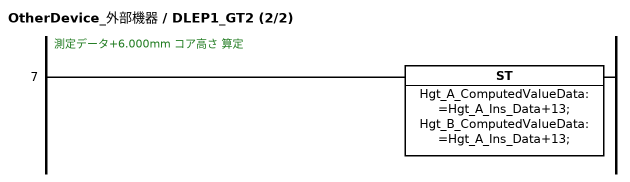
(* [picture p96: OtherDevice_外部機器 / DLEP1_GT2, rungs 7-7] *)
(* Rung 7: 測定データ+6.000mm コア高さ 算定 *)
Hgt_A_ComputedValueData:=Hgt_A_Ins_Data+13;
Hgt_B_ComputedValueData:=Hgt_A_Ins_Data+13;

(* Section FH_5552_10: ladder, written here as Structured Text *)

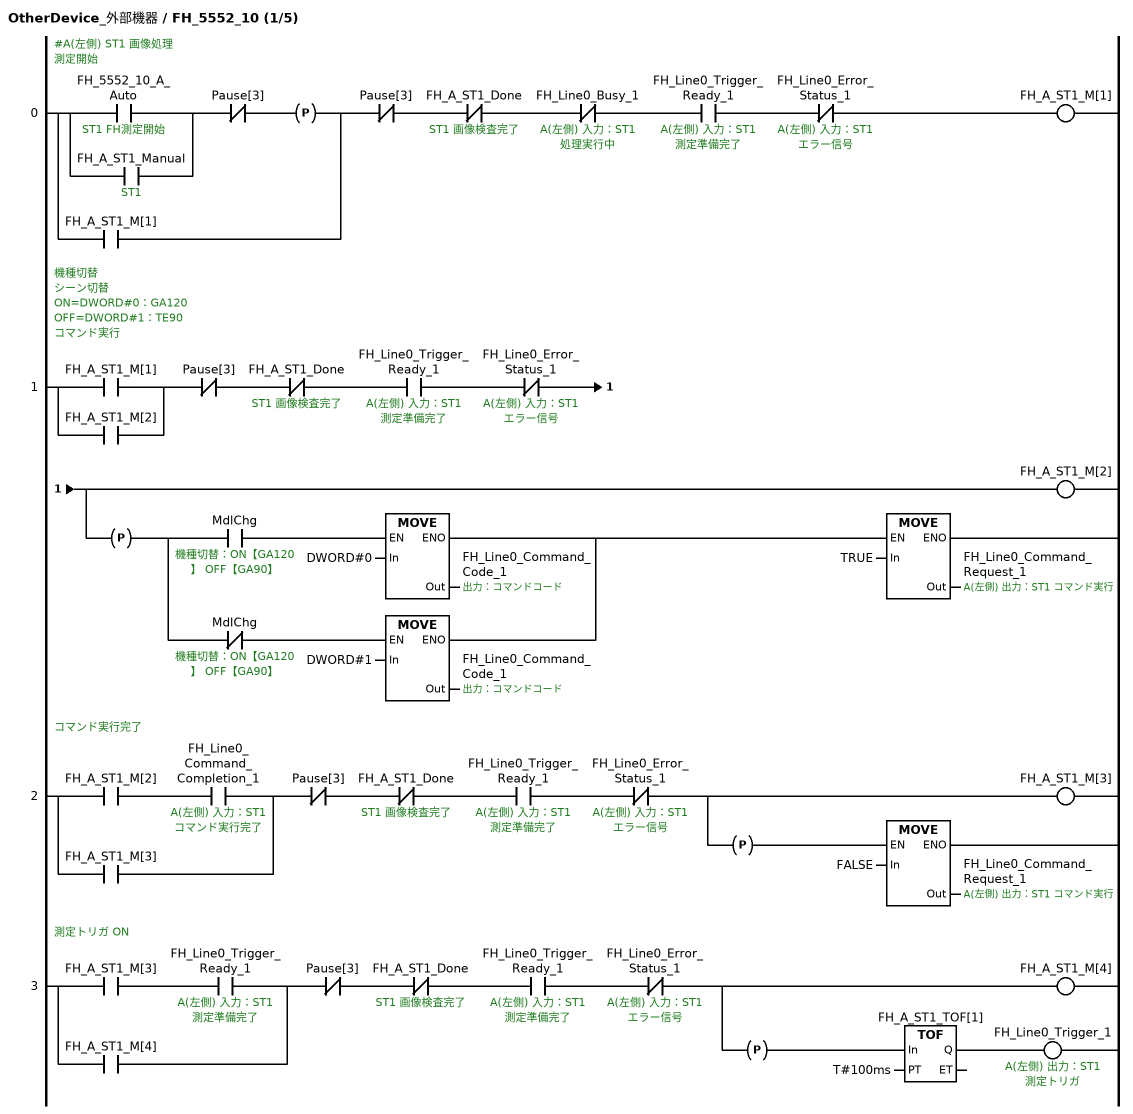
(* Rung 0: #A(左側) ST1 画像処理 / 測定開始 *)
_e25(CLK := (FH_5552_10_A_Auto OR FH_A_ST1_Manual) AND NOT Pause[3]);
FH_A_ST1_M[1] := (_e25.Q OR FH_A_ST1_M[1]) AND NOT Pause[3] AND NOT FH_A_ST1_Done AND NOT FH_Line0_Busy_1 AND FH_Line0_Trigger_Ready_1 AND NOT FH_Line0_Error_Status_1;
(* Rung 1: 機種切替 / シーン切替 / ON=DWORD#0：GA120 / OFF=DWORD#1：TE90 / コマンド実行 *)
_p26 := (FH_A_ST1_M[1] OR FH_A_ST1_M[2]) AND NOT Pause[3] AND NOT FH_A_ST1_Done AND FH_Line0_Trigger_Ready_1 AND NOT FH_Line0_Error_Status_1;
FH_A_ST1_M[2] := _p26;
_e27(CLK := _p26);
IF _e27.Q AND MdlChg THEN FH_Line0_Command_Code_1 := DWORD#0; END_IF;
IF _e27.Q AND NOT MdlChg THEN FH_Line0_Command_Code_1 := DWORD#1; END_IF;
IF _e27.Q AND (MdlChg OR NOT MdlChg) THEN FH_Line0_Command_Request_1 := TRUE; END_IF;
(* Rung 2: コマンド実行完了 *)
_p28 := ((FH_A_ST1_M[2] AND FH_Line0_Command_Completion_1) OR FH_A_ST1_M[3]) AND NOT Pause[3] AND NOT FH_A_ST1_Done AND FH_Line0_Trigger_Ready_1 AND NOT FH_Line0_Error_Status_1;
FH_A_ST1_M[3] := _p28;
_e29(CLK := _p28);
IF _e29.Q THEN FH_Line0_Command_Request_1 := FALSE; END_IF;
(* Rung 3: 測定トリガ ON *)
_p30 := ((FH_A_ST1_M[3] AND FH_Line0_Trigger_Ready_1) OR FH_A_ST1_M[4]) AND NOT Pause[3] AND NOT FH_A_ST1_Done AND FH_Line0_Trigger_Ready_1 AND NOT FH_Line0_Error_Status_1;
FH_A_ST1_M[4] := _p30;
_e31(CLK := _p30);
FH_A_ST1_TOF[1](In := _e31.Q, PT := T#100ms);
FH_Line0_Trigger_1 := FH_A_ST1_TOF[1].Q;

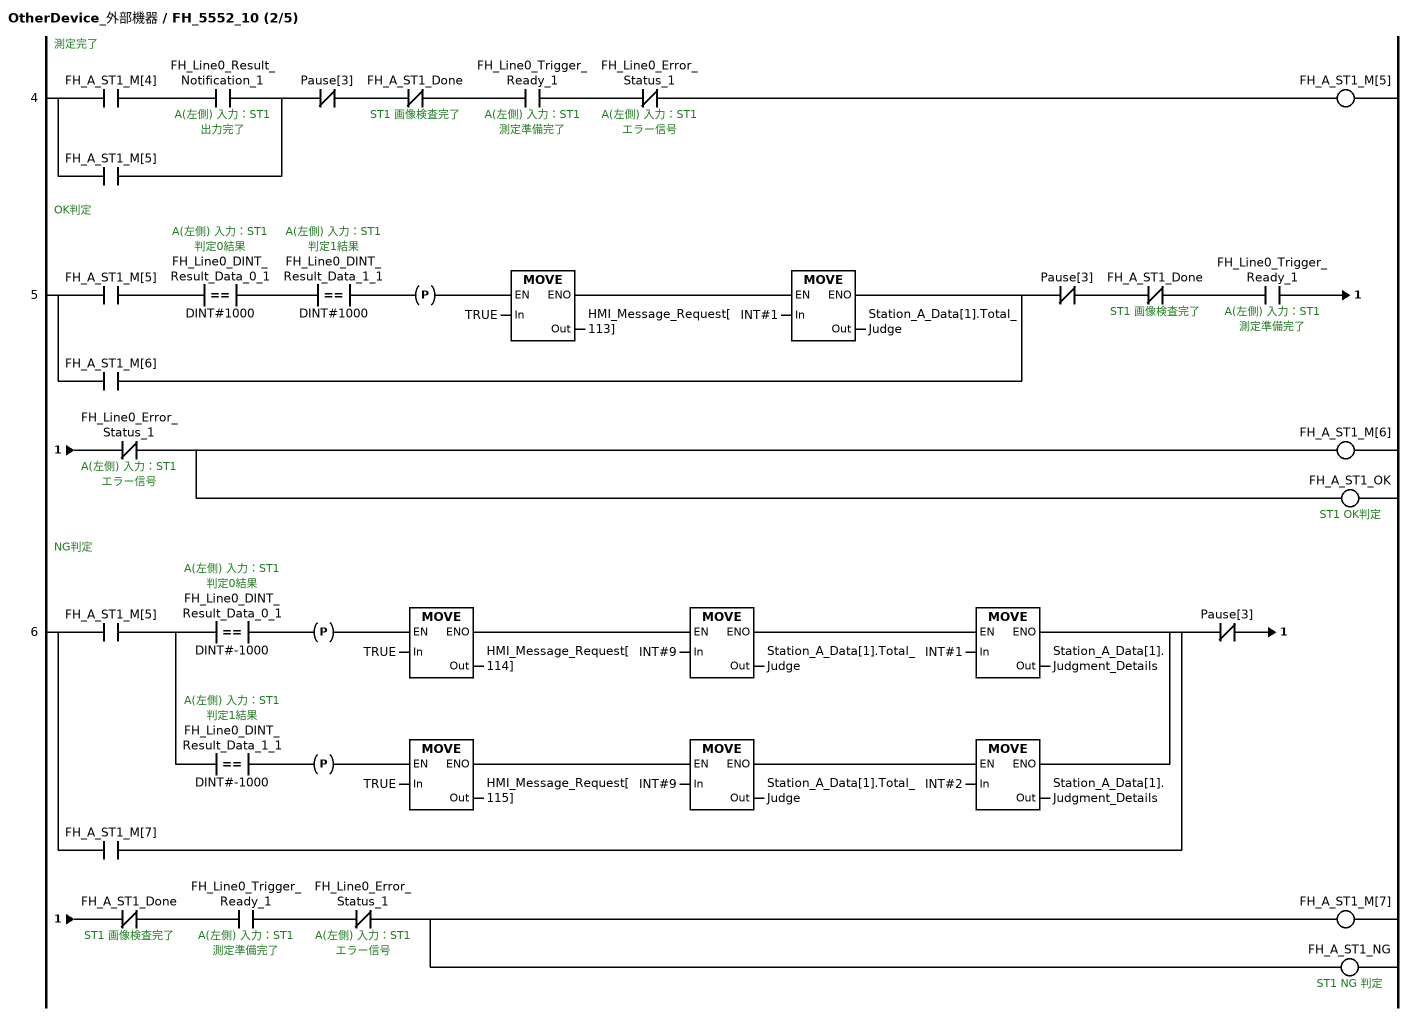
(* Rung 4: 測定完了 *)
FH_A_ST1_M[5] := ((FH_A_ST1_M[4] AND FH_Line0_Result_Notification_1) OR FH_A_ST1_M[5]) AND NOT Pause[3] AND NOT FH_A_ST1_Done AND FH_Line0_Trigger_Ready_1 AND NOT FH_Line0_Error_Status_1;
(* Rung 5: OK判定 *)
_e32(CLK := FH_A_ST1_M[5] AND (FH_Line0_DINT_Result_Data_0_1 = DINT#1000) AND (FH_Line0_DINT_Result_Data_1_1 = DINT#1000));
IF _e32.Q THEN
    HMI_Message_Request[113] := TRUE;
    Station_A_Data[1].Total_Judge := INT#1;
END_IF;
_p33 := (_e32.Q OR FH_A_ST1_M[6]) AND NOT Pause[3] AND NOT FH_A_ST1_Done AND FH_Line0_Trigger_Ready_1 AND NOT FH_Line0_Error_Status_1;
FH_A_ST1_M[6] := _p33;
FH_A_ST1_OK := _p33;
(* Rung 6: NG判定 *)
_e34(CLK := FH_A_ST1_M[5] AND (FH_Line0_DINT_Result_Data_0_1 = (DINT#-1000)));
IF _e34.Q THEN
    HMI_Message_Request[114] := TRUE;
    Station_A_Data[1].Total_Judge := INT#9;
    Station_A_Data[1].Judgment_Details := INT#1;
END_IF;
_e35(CLK := FH_A_ST1_M[5] AND (FH_Line0_DINT_Result_Data_1_1 = (DINT#-1000)));
IF _e35.Q THEN
    HMI_Message_Request[115] := TRUE;
    Station_A_Data[1].Total_Judge := INT#9;
    Station_A_Data[1].Judgment_Details := INT#2;
END_IF;
_p36 := (_e34.Q OR _e35.Q OR FH_A_ST1_M[7]) AND NOT Pause[3] AND NOT FH_A_ST1_Done AND FH_Line0_Trigger_Ready_1 AND NOT FH_Line0_Error_Status_1;
FH_A_ST1_M[7] := _p36;
FH_A_ST1_NG := _p36;

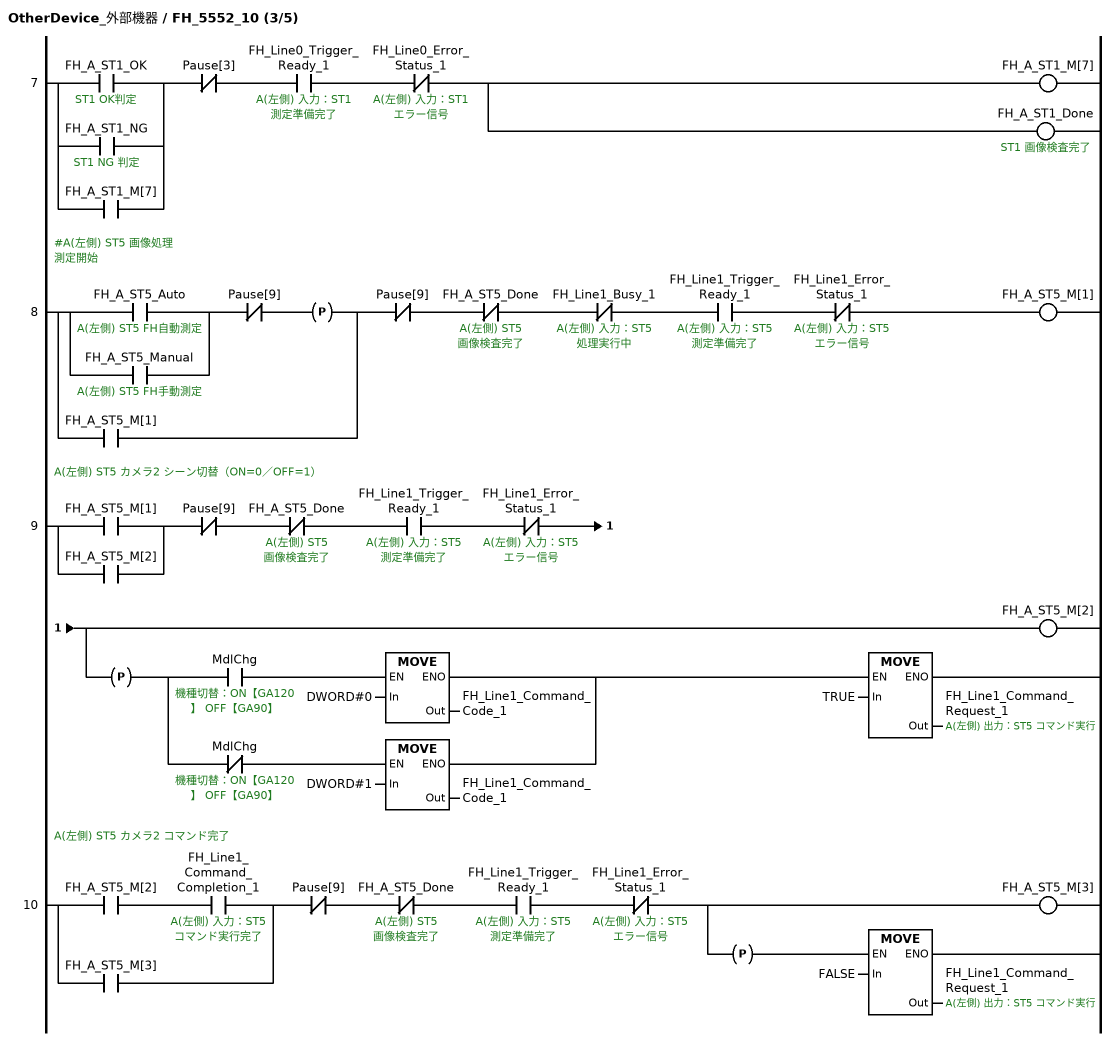
(* Rung 7 *)
_p37 := (FH_A_ST1_OK OR FH_A_ST1_NG OR FH_A_ST1_M[7]) AND NOT Pause[3] AND FH_Line0_Trigger_Ready_1 AND NOT FH_Line0_Error_Status_1;
FH_A_ST1_M[7] := _p37;
FH_A_ST1_Done := _p37;
(* Rung 8: #A(左側) ST5 画像処理 / 測定開始 *)
_e38(CLK := (FH_A_ST5_Auto OR FH_A_ST5_Manual) AND NOT Pause[9]);
FH_A_ST5_M[1] := (_e38.Q OR FH_A_ST5_M[1]) AND NOT Pause[9] AND NOT FH_A_ST5_Done AND NOT FH_Line1_Busy_1 AND FH_Line1_Trigger_Ready_1 AND NOT FH_Line1_Error_Status_1;
(* Rung 9: A(左側) ST5 カメラ2 シーン切替（ON=0／OFF=1） *)
_p39 := (FH_A_ST5_M[1] OR FH_A_ST5_M[2]) AND NOT Pause[9] AND NOT FH_A_ST5_Done AND FH_Line1_Trigger_Ready_1 AND NOT FH_Line1_Error_Status_1;
FH_A_ST5_M[2] := _p39;
_e40(CLK := _p39);
IF _e40.Q AND MdlChg THEN FH_Line1_Command_Code_1 := DWORD#0; END_IF;
IF _e40.Q AND NOT MdlChg THEN FH_Line1_Command_Code_1 := DWORD#1; END_IF;
IF _e40.Q AND (MdlChg OR NOT MdlChg) THEN FH_Line1_Command_Request_1 := TRUE; END_IF;
(* Rung 10: A(左側) ST5 カメラ2 コマンド完了 *)
_p41 := ((FH_A_ST5_M[2] AND FH_Line1_Command_Completion_1) OR FH_A_ST5_M[3]) AND NOT Pause[9] AND NOT FH_A_ST5_Done AND FH_Line1_Trigger_Ready_1 AND NOT FH_Line1_Error_Status_1;
FH_A_ST5_M[3] := _p41;
_e42(CLK := _p41);
IF _e42.Q THEN FH_Line1_Command_Request_1 := FALSE; END_IF;

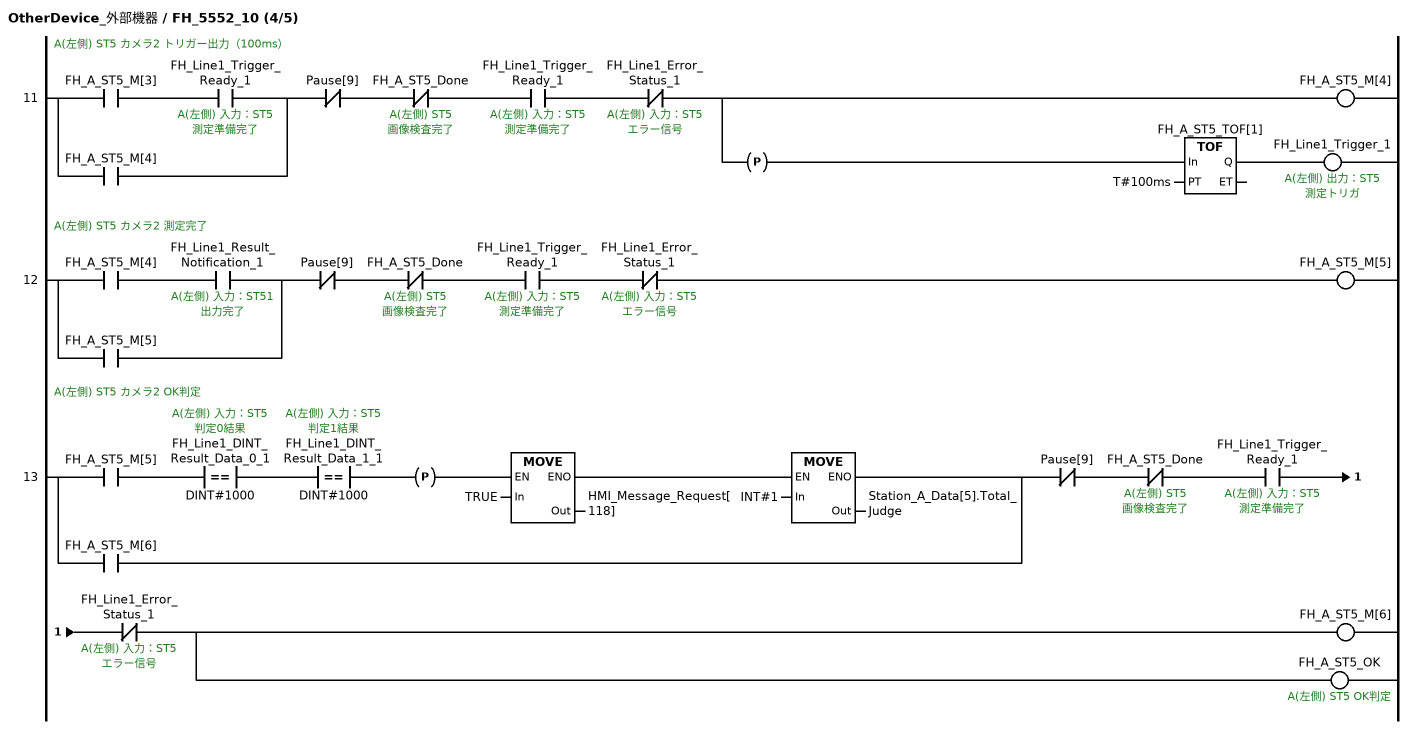
(* Rung 11: A(左側) ST5 カメラ2 トリガー出力（100ms） *)
_p43 := ((FH_A_ST5_M[3] AND FH_Line1_Trigger_Ready_1) OR FH_A_ST5_M[4]) AND NOT Pause[9] AND NOT FH_A_ST5_Done AND FH_Line1_Trigger_Ready_1 AND NOT FH_Line1_Error_Status_1;
FH_A_ST5_M[4] := _p43;
_e44(CLK := _p43);
FH_A_ST5_TOF[1](In := _e44.Q, PT := T#100ms);
FH_Line1_Trigger_1 := FH_A_ST5_TOF[1].Q;
(* Rung 12: A(左側) ST5 カメラ2 測定完了 *)
FH_A_ST5_M[5] := ((FH_A_ST5_M[4] AND FH_Line1_Result_Notification_1) OR FH_A_ST5_M[5]) AND NOT Pause[9] AND NOT FH_A_ST5_Done AND FH_Line1_Trigger_Ready_1 AND NOT FH_Line1_Error_Status_1;
(* Rung 13: A(左側) ST5 カメラ2 OK判定 *)
_e45(CLK := FH_A_ST5_M[5] AND (FH_Line1_DINT_Result_Data_0_1 = DINT#1000) AND (FH_Line1_DINT_Result_Data_1_1 = DINT#1000));
IF _e45.Q THEN
    HMI_Message_Request[118] := TRUE;
    Station_A_Data[5].Total_Judge := INT#1;
END_IF;
_p46 := (_e45.Q OR FH_A_ST5_M[6]) AND NOT Pause[9] AND NOT FH_A_ST5_Done AND FH_Line1_Trigger_Ready_1 AND NOT FH_Line1_Error_Status_1;
FH_A_ST5_M[6] := _p46;
FH_A_ST5_OK := _p46;

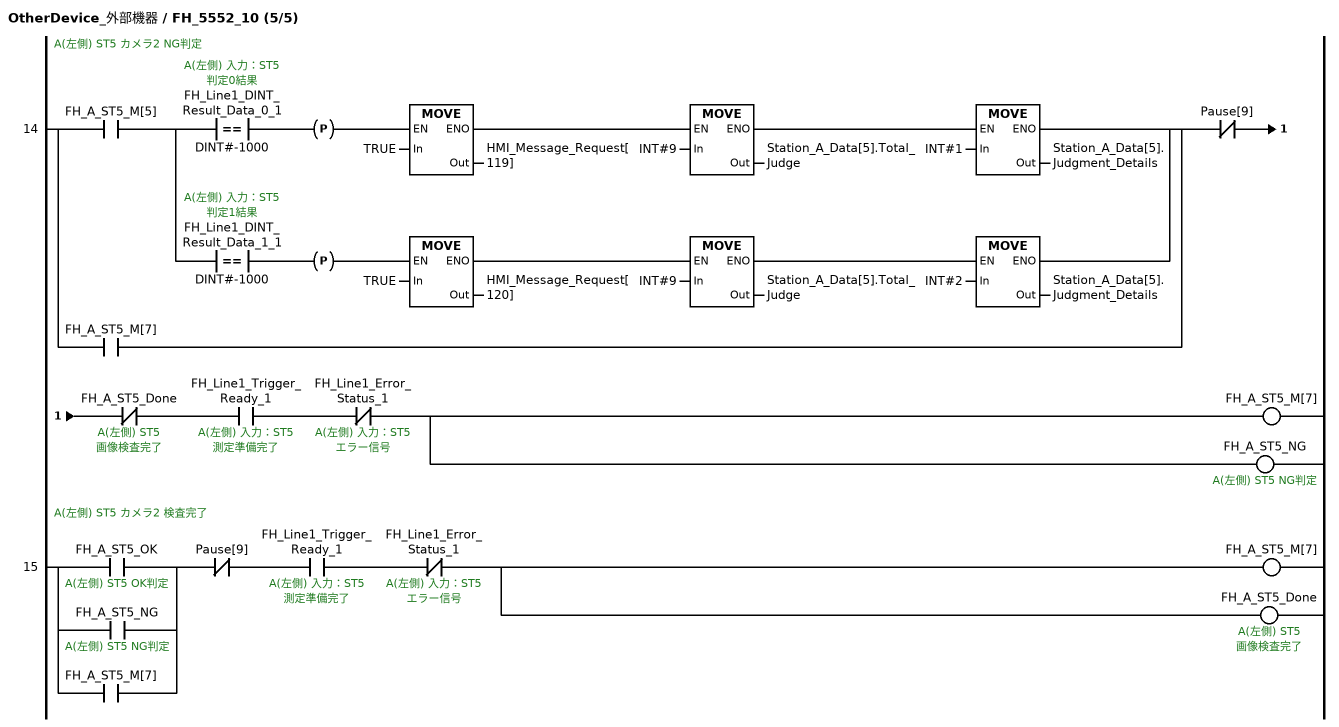
(* Rung 14: A(左側) ST5 カメラ2 NG判定 *)
_e47(CLK := FH_A_ST5_M[5] AND (FH_Line1_DINT_Result_Data_0_1 = (DINT#-1000)));
IF _e47.Q THEN
    HMI_Message_Request[119] := TRUE;
    Station_A_Data[5].Total_Judge := INT#9;
    Station_A_Data[5].Judgment_Details := INT#1;
END_IF;
_e48(CLK := FH_A_ST5_M[5] AND (FH_Line1_DINT_Result_Data_1_1 = (DINT#-1000)));
IF _e48.Q THEN
    HMI_Message_Request[120] := TRUE;
    Station_A_Data[5].Total_Judge := INT#9;
    Station_A_Data[5].Judgment_Details := INT#2;
END_IF;
_p49 := (_e47.Q OR _e48.Q OR FH_A_ST5_M[7]) AND NOT Pause[9] AND NOT FH_A_ST5_Done AND FH_Line1_Trigger_Ready_1 AND NOT FH_Line1_Error_Status_1;
FH_A_ST5_M[7] := _p49;
FH_A_ST5_NG := _p49;
(* Rung 15: A(左側) ST5 カメラ2 検査完了 *)
_p50 := (FH_A_ST5_OK OR FH_A_ST5_NG OR FH_A_ST5_M[7]) AND NOT Pause[9] AND FH_Line1_Trigger_Ready_1 AND NOT FH_Line1_Error_Status_1;
FH_A_ST5_M[7] := _p50;
FH_A_ST5_Done := _p50;

(* Section CV2A_KED: ladder, written here as Structured Text *)

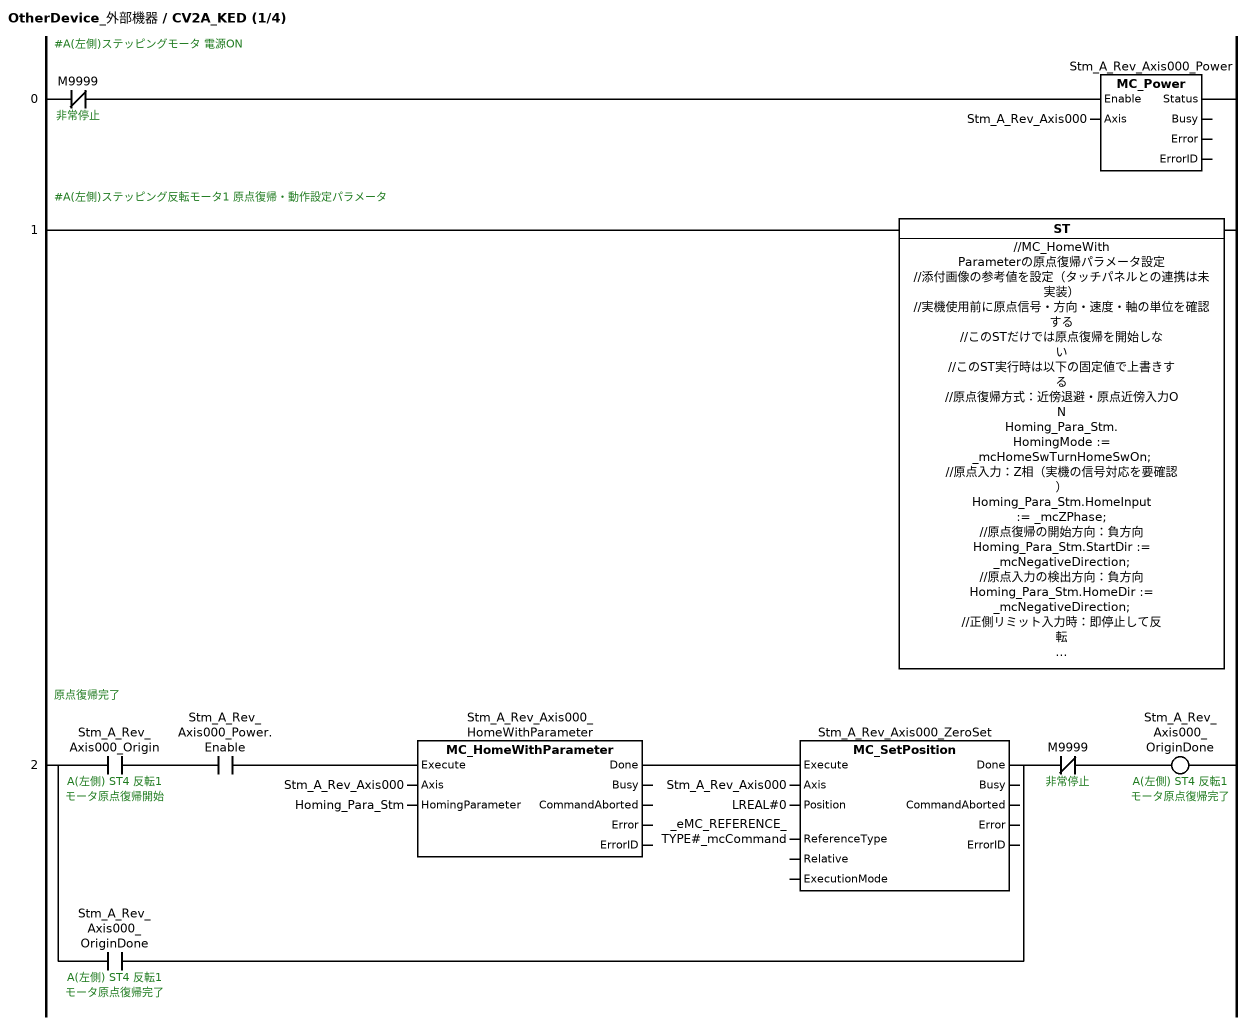
(* Rung 0: #A(左側)ステッピングモータ 電源ON *)
Stm_A_Rev_Axis000_Power(Enable := NOT M9999, Axis := Stm_A_Rev_Axis000);
(* Rung 1: #A(左側)ステッピング反転モータ1 原点復帰・動作設定パラメータ *)
//MC_HomeWithParameterの原点復帰パラメータ設定
//添付画像の参考値を設定（タッチパネルとの連携は未実装）
//実機使用前に原点信号・方向・速度・軸の単位を確認する
//このSTだけでは原点復帰を開始しない
//このST実行時は以下の固定値で上書きする

//原点復帰方式：近傍退避・原点近傍入力ON
Homing_Para_Stm.HomingMode := _mcHomeSwTurnHomeSwOn;
//原点入力：Z相（実機の信号対応を要確認）
Homing_Para_Stm.HomeInput := _mcZPhase;
//原点復帰の開始方向：負方向
Homing_Para_Stm.StartDir := _mcNegativeDirection;
//原点入力の検出方向：負方向
Homing_Para_Stm.HomeDir := _mcNegativeDirection;
//正側リミット入力時：即停止して反転
Homing_Para_Stm.PosiLmtMode := _mcRevImmediateStop;
//負側リミット入力時：即停止して反転
Homing_Para_Stm.NegaLmtMode := _mcRevImmediateStop;

//原点復帰速度 [指令単位/s]
Homing_Para_Stm.Vel := LREAL#40;
//原点近傍での接近速度 [指令単位/s]
Homing_Para_Stm.ApproachVel := LREAL#1;
//原点復帰の加速度 [指令単位/s^2]
Homing_Para_Stm.Acc := LREAL#100;
//原点復帰の減速度 [指令単位/s^2]
Homing_Para_Stm.Dec := LREAL#200;
//ジャーク [指令単位/s^3]：0はジャーク制御なし
Homing_Para_Stm.Jerk := LREAL#0;

//原点入力マスク距離 [指令単位]：今回の方式では未使用
Homing_Para_Stm.Mask := LREAL#0;
//原点確定後の現在位置 [指令単位]
Homing_Para_Stm.Offset := LREAL#0;
//押当て時間 [ms]：今回の方式では未使用
Homing_Para_Stm.PushTime := UINT#0;
//原点検出後の補正移動量 [指令単位]：0は補正移動なし
Homing_Para_Stm.Compensation := LREAL#0;
//原点補正移動時の速度 [指令単位/s]
Homing_Para_Stm.CompensationVel := LREAL#10;
(* Rung 2: 原点復帰完了 *)
Stm_A_Rev_Axis000_HomeWithParameter(Execute := Stm_A_Rev_Axis000_Origin AND Stm_A_Rev_Axis000_Power.Enable, Axis := Stm_A_Rev_Axis000, HomingParameter := Homing_Para_Stm);
Stm_A_Rev_Axis000_ZeroSet(Execute := Stm_A_Rev_Axis000_HomeWithParameter.Done, Axis := Stm_A_Rev_Axis000, Position := LREAL#0, ReferenceType := _eMC_REFERENCE_TYPE#_mcCommand);
Stm_A_Rev_Axis000_OriginDone := (Stm_A_Rev_Axis000_ZeroSet.Done OR Stm_A_Rev_Axis000_OriginDone) AND NOT M9999;

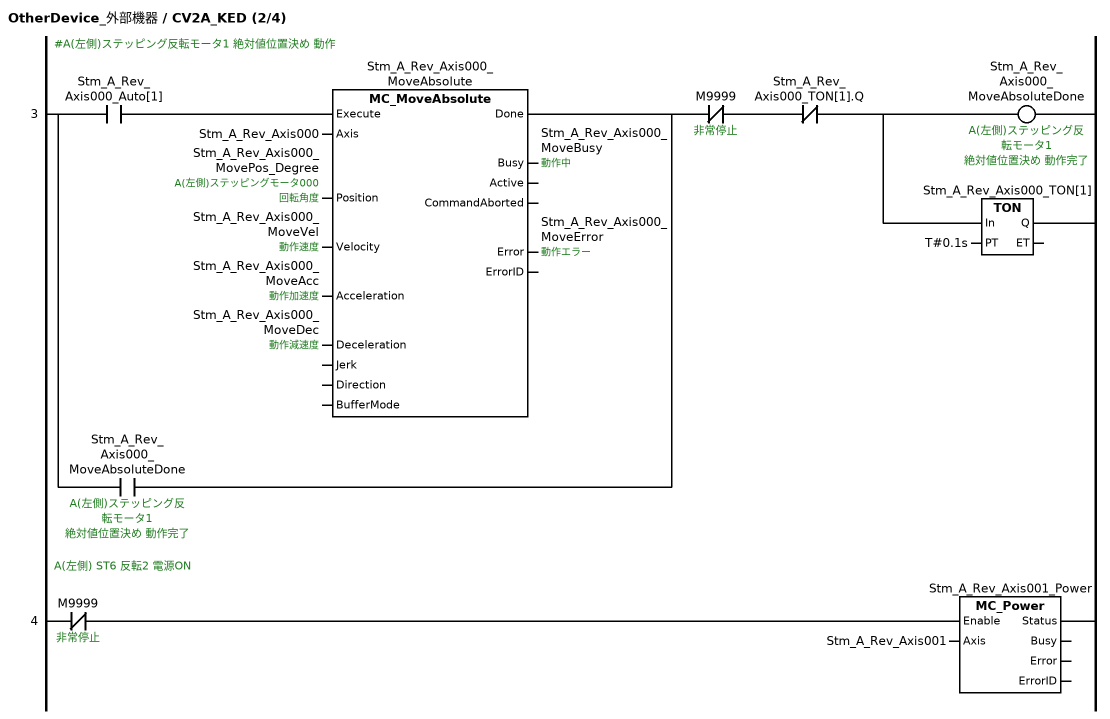
(* Rung 3: #A(左側)ステッピング反転モータ1 絶対値位置決め 動作 *)
Stm_A_Rev_Axis000_MoveAbsolute(Execute := Stm_A_Rev_Axis000_Auto[1], Axis := Stm_A_Rev_Axis000, Position := Stm_A_Rev_Axis000_MovePos_Degree, Velocity := Stm_A_Rev_Axis000_MoveVel, Acceleration := Stm_A_Rev_Axis000_MoveAcc, Deceleration := Stm_A_Rev_Axis000_MoveDec, Busy => Stm_A_Rev_Axis000_MoveBusy, Error => Stm_A_Rev_Axis000_MoveError);
_p51 := (Stm_A_Rev_Axis000_MoveAbsolute.Done OR Stm_A_Rev_Axis000_MoveAbsoluteDone) AND NOT M9999 AND NOT Stm_A_Rev_Axis000_TON[1].Q;
Stm_A_Rev_Axis000_MoveAbsoluteDone := _p51;
Stm_A_Rev_Axis000_TON[1](In := _p51, PT := T#0.1s);
(* Rung 4: A(左側) ST6 反転2 電源ON *)
Stm_A_Rev_Axis001_Power(Enable := NOT M9999, Axis := Stm_A_Rev_Axis001);

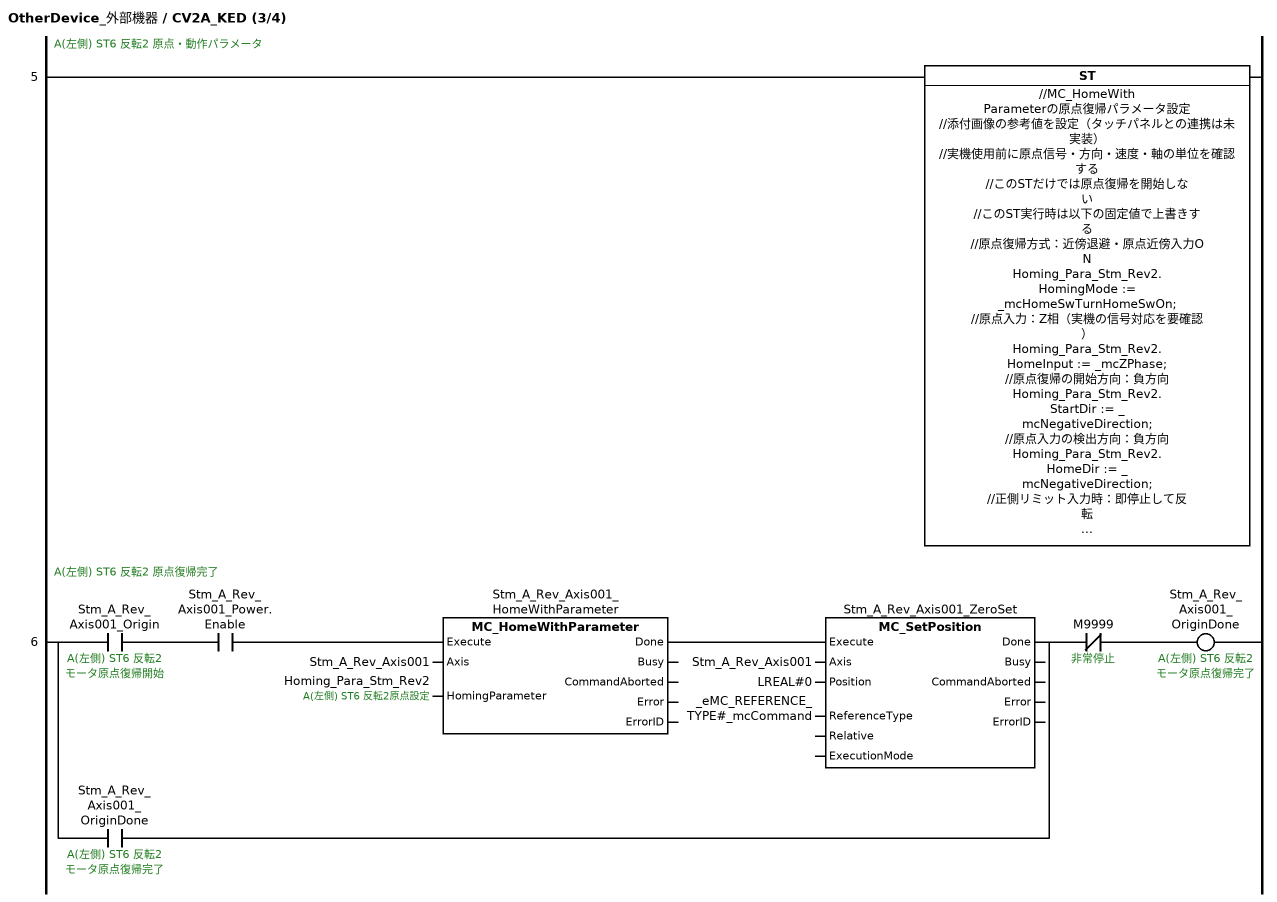
(* Rung 5: A(左側) ST6 反転2 原点・動作パラメータ *)
//MC_HomeWithParameterの原点復帰パラメータ設定
//添付画像の参考値を設定（タッチパネルとの連携は未実装）
//実機使用前に原点信号・方向・速度・軸の単位を確認する
//このSTだけでは原点復帰を開始しない
//このST実行時は以下の固定値で上書きする

//原点復帰方式：近傍退避・原点近傍入力ON
Homing_Para_Stm_Rev2.HomingMode := _mcHomeSwTurnHomeSwOn;
//原点入力：Z相（実機の信号対応を要確認）
Homing_Para_Stm_Rev2.HomeInput := _mcZPhase;
//原点復帰の開始方向：負方向
Homing_Para_Stm_Rev2.StartDir := _mcNegativeDirection;
//原点入力の検出方向：負方向
Homing_Para_Stm_Rev2.HomeDir := _mcNegativeDirection;
//正側リミット入力時：即停止して反転
Homing_Para_Stm_Rev2.PosiLmtMode := _mcRevImmediateStop;
//負側リミット入力時：即停止して反転
Homing_Para_Stm_Rev2.NegaLmtMode := _mcRevImmediateStop;

//原点復帰速度 [指令単位/s]
Homing_Para_Stm_Rev2.Vel := LREAL#40;
//原点近傍での接近速度 [指令単位/s]
Homing_Para_Stm_Rev2.ApproachVel := LREAL#1;
//原点復帰の加速度 [指令単位/s^2]
Homing_Para_Stm_Rev2.Acc := LREAL#100;
//原点復帰の減速度 [指令単位/s^2]
Homing_Para_Stm_Rev2.Dec := LREAL#200;
//ジャーク [指令単位/s^3]：0はジャーク制御なし
Homing_Para_Stm_Rev2.Jerk := LREAL#0;

//原点入力マスク距離 [指令単位]：今回の方式では未使用
Homing_Para_Stm_Rev2.Mask := LREAL#0;
//原点確定後の現在位置 [指令単位]
Homing_Para_Stm_Rev2.Offset := LREAL#0;
//押当て時間 [ms]：今回の方式では未使用
Homing_Para_Stm_Rev2.PushTime := UINT#0;
//原点検出後の補正移動量 [指令単位]：0は補正移動なし
Homing_Para_Stm_Rev2.Compensation := LREAL#0;
//原点補正移動時の速度 [指令単位/s]
Homing_Para_Stm_Rev2.CompensationVel := LREAL#10;
(* Rung 6: A(左側) ST6 反転2 原点復帰完了 *)
Stm_A_Rev_Axis001_HomeWithParameter(Execute := Stm_A_Rev_Axis001_Origin AND Stm_A_Rev_Axis001_Power.Enable, Axis := Stm_A_Rev_Axis001, HomingParameter := Homing_Para_Stm_Rev2);
Stm_A_Rev_Axis001_ZeroSet(Execute := Stm_A_Rev_Axis001_HomeWithParameter.Done, Axis := Stm_A_Rev_Axis001, Position := LREAL#0, ReferenceType := _eMC_REFERENCE_TYPE#_mcCommand);
Stm_A_Rev_Axis001_OriginDone := (Stm_A_Rev_Axis001_ZeroSet.Done OR Stm_A_Rev_Axis001_OriginDone) AND NOT M9999;

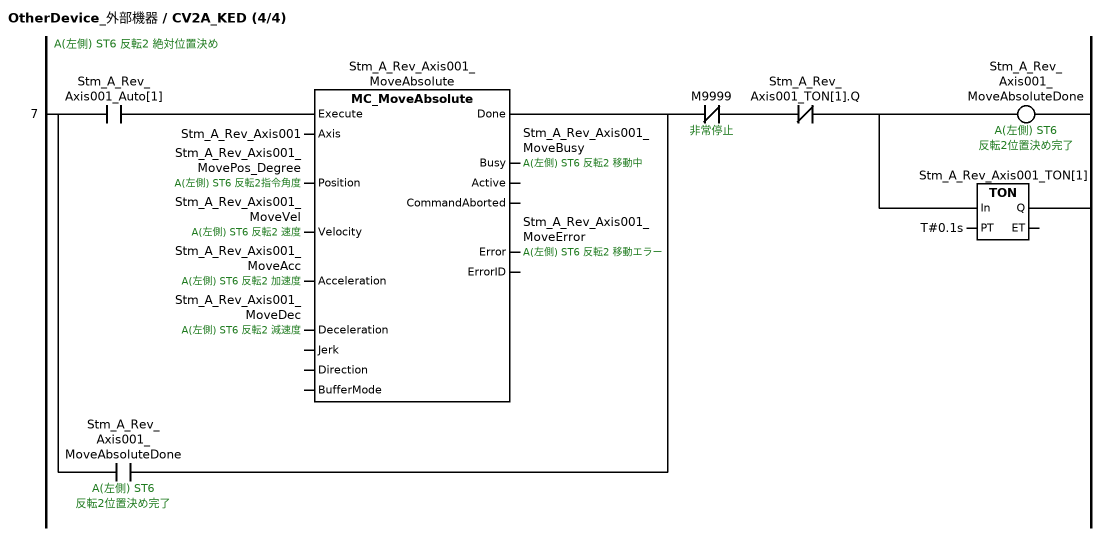
(* Rung 7: A(左側) ST6 反転2 絶対位置決め *)
Stm_A_Rev_Axis001_MoveAbsolute(Execute := Stm_A_Rev_Axis001_Auto[1], Axis := Stm_A_Rev_Axis001, Position := Stm_A_Rev_Axis001_MovePos_Degree, Velocity := Stm_A_Rev_Axis001_MoveVel, Acceleration := Stm_A_Rev_Axis001_MoveAcc, Deceleration := Stm_A_Rev_Axis001_MoveDec, Busy => Stm_A_Rev_Axis001_MoveBusy, Error => Stm_A_Rev_Axis001_MoveError);
_p52 := (Stm_A_Rev_Axis001_MoveAbsolute.Done OR Stm_A_Rev_Axis001_MoveAbsoluteDone) AND NOT M9999 AND NOT Stm_A_Rev_Axis001_TON[1].Q;
Stm_A_Rev_Axis001_MoveAbsoluteDone := _p52;
Stm_A_Rev_Axis001_TON[1](In := _p52, PT := T#0.1s);

(* Section HMI: ladder, written here as Structured Text *)

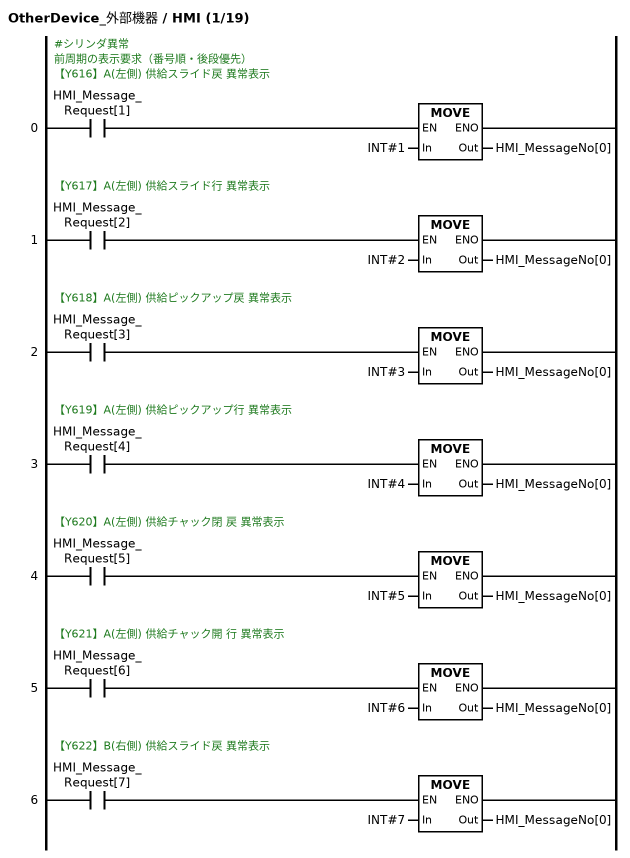
(* Rung 0: #シリンダ異常 / 前周期の表示要求（番号順・後段優先） / 【Y616】A(左側) 供給スライド戻 異常表示 *)
IF HMI_Message_Request[1] THEN HMI_MessageNo[0] := INT#1; END_IF;
(* Rung 1: 【Y617】A(左側) 供給スライド行 異常表示 *)
IF HMI_Message_Request[2] THEN HMI_MessageNo[0] := INT#2; END_IF;
(* Rung 2: 【Y618】A(左側) 供給ピックアップ戻 異常表示 *)
IF HMI_Message_Request[3] THEN HMI_MessageNo[0] := INT#3; END_IF;
(* Rung 3: 【Y619】A(左側) 供給ピックアップ行 異常表示 *)
IF HMI_Message_Request[4] THEN HMI_MessageNo[0] := INT#4; END_IF;
(* Rung 4: 【Y620】A(左側) 供給チャック閉 戻 異常表示 *)
IF HMI_Message_Request[5] THEN HMI_MessageNo[0] := INT#5; END_IF;
(* Rung 5: 【Y621】A(左側) 供給チャック開 行 異常表示 *)
IF HMI_Message_Request[6] THEN HMI_MessageNo[0] := INT#6; END_IF;
(* Rung 6: 【Y622】B(右側) 供給スライド戻 異常表示 *)
IF HMI_Message_Request[7] THEN HMI_MessageNo[0] := INT#7; END_IF;

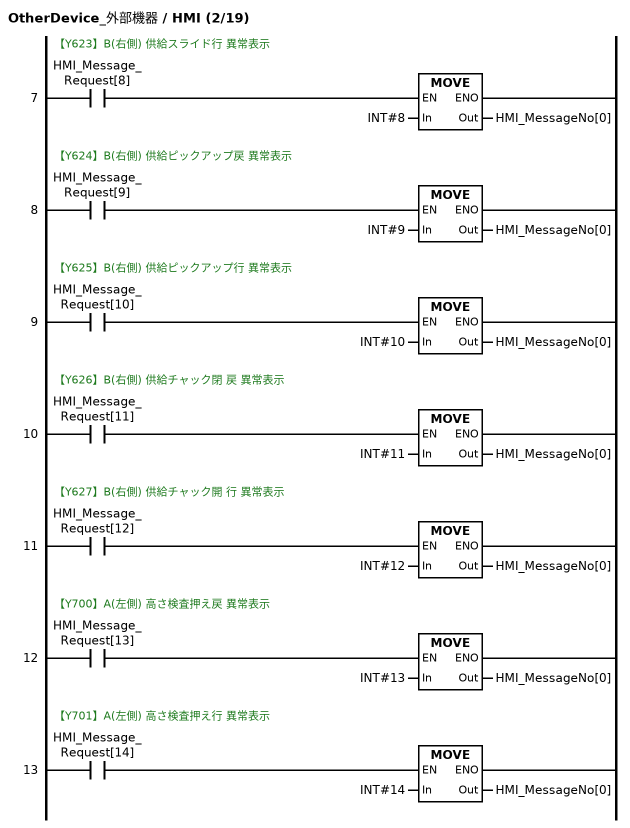
(* Rung 7: 【Y623】B(右側) 供給スライド行 異常表示 *)
IF HMI_Message_Request[8] THEN HMI_MessageNo[0] := INT#8; END_IF;
(* Rung 8: 【Y624】B(右側) 供給ピックアップ戻 異常表示 *)
IF HMI_Message_Request[9] THEN HMI_MessageNo[0] := INT#9; END_IF;
(* Rung 9: 【Y625】B(右側) 供給ピックアップ行 異常表示 *)
IF HMI_Message_Request[10] THEN HMI_MessageNo[0] := INT#10; END_IF;
(* Rung 10: 【Y626】B(右側) 供給チャック閉 戻 異常表示 *)
IF HMI_Message_Request[11] THEN HMI_MessageNo[0] := INT#11; END_IF;
(* Rung 11: 【Y627】B(右側) 供給チャック開 行 異常表示 *)
IF HMI_Message_Request[12] THEN HMI_MessageNo[0] := INT#12; END_IF;
(* Rung 12: 【Y700】A(左側) 高さ検査押え戻 異常表示 *)
IF HMI_Message_Request[13] THEN HMI_MessageNo[0] := INT#13; END_IF;
(* Rung 13: 【Y701】A(左側) 高さ検査押え行 異常表示 *)
IF HMI_Message_Request[14] THEN HMI_MessageNo[0] := INT#14; END_IF;

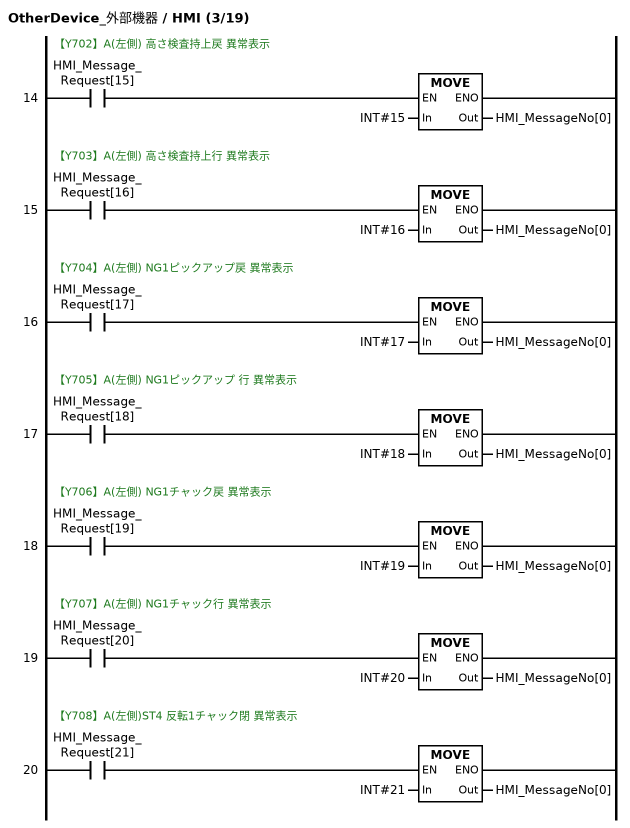
(* Rung 14: 【Y702】A(左側) 高さ検査持上戻 異常表示 *)
IF HMI_Message_Request[15] THEN HMI_MessageNo[0] := INT#15; END_IF;
(* Rung 15: 【Y703】A(左側) 高さ検査持上行 異常表示 *)
IF HMI_Message_Request[16] THEN HMI_MessageNo[0] := INT#16; END_IF;
(* Rung 16: 【Y704】A(左側) NG1ピックアップ戻 異常表示 *)
IF HMI_Message_Request[17] THEN HMI_MessageNo[0] := INT#17; END_IF;
(* Rung 17: 【Y705】A(左側) NG1ピックアップ 行 異常表示 *)
IF HMI_Message_Request[18] THEN HMI_MessageNo[0] := INT#18; END_IF;
(* Rung 18: 【Y706】A(左側) NG1チャック戻 異常表示 *)
IF HMI_Message_Request[19] THEN HMI_MessageNo[0] := INT#19; END_IF;
(* Rung 19: 【Y707】A(左側) NG1チャック行 異常表示 *)
IF HMI_Message_Request[20] THEN HMI_MessageNo[0] := INT#20; END_IF;
(* Rung 20: 【Y708】A(左側)ST4 反転1チャック閉 異常表示 *)
IF HMI_Message_Request[21] THEN HMI_MessageNo[0] := INT#21; END_IF;

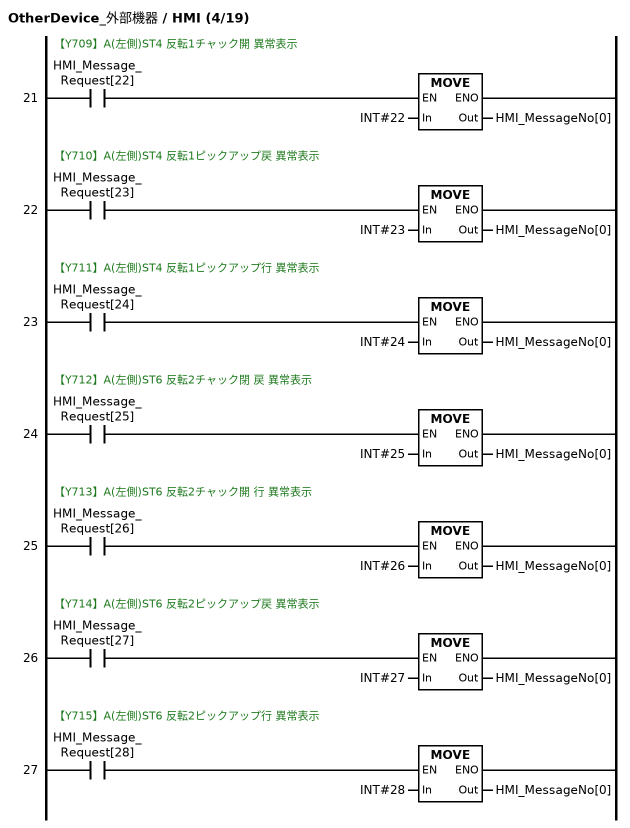
(* Rung 21: 【Y709】A(左側)ST4 反転1チャック開 異常表示 *)
IF HMI_Message_Request[22] THEN HMI_MessageNo[0] := INT#22; END_IF;
(* Rung 22: 【Y710】A(左側)ST4 反転1ピックアップ戻 異常表示 *)
IF HMI_Message_Request[23] THEN HMI_MessageNo[0] := INT#23; END_IF;
(* Rung 23: 【Y711】A(左側)ST4 反転1ピックアップ行 異常表示 *)
IF HMI_Message_Request[24] THEN HMI_MessageNo[0] := INT#24; END_IF;
(* Rung 24: 【Y712】A(左側)ST6 反転2チャック閉 戻 異常表示 *)
IF HMI_Message_Request[25] THEN HMI_MessageNo[0] := INT#25; END_IF;
(* Rung 25: 【Y713】A(左側)ST6 反転2チャック開 行 異常表示 *)
IF HMI_Message_Request[26] THEN HMI_MessageNo[0] := INT#26; END_IF;
(* Rung 26: 【Y714】A(左側)ST6 反転2ピックアップ戻 異常表示 *)
IF HMI_Message_Request[27] THEN HMI_MessageNo[0] := INT#27; END_IF;
(* Rung 27: 【Y715】A(左側)ST6 反転2ピックアップ行 異常表示 *)
IF HMI_Message_Request[28] THEN HMI_MessageNo[0] := INT#28; END_IF;

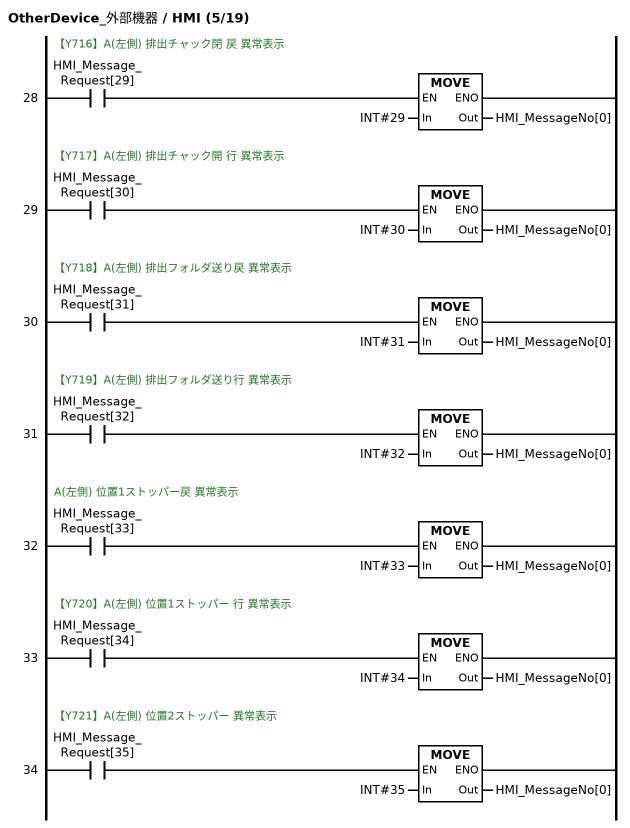
(* Rung 28: 【Y716】A(左側) 排出チャック閉 戻 異常表示 *)
IF HMI_Message_Request[29] THEN HMI_MessageNo[0] := INT#29; END_IF;
(* Rung 29: 【Y717】A(左側) 排出チャック開 行 異常表示 *)
IF HMI_Message_Request[30] THEN HMI_MessageNo[0] := INT#30; END_IF;
(* Rung 30: 【Y718】A(左側) 排出フォルダ送り戻 異常表示 *)
IF HMI_Message_Request[31] THEN HMI_MessageNo[0] := INT#31; END_IF;
(* Rung 31: 【Y719】A(左側) 排出フォルダ送り行 異常表示 *)
IF HMI_Message_Request[32] THEN HMI_MessageNo[0] := INT#32; END_IF;
(* Rung 32: A(左側) 位置1ストッパー戻 異常表示 *)
IF HMI_Message_Request[33] THEN HMI_MessageNo[0] := INT#33; END_IF;
(* Rung 33: 【Y720】A(左側) 位置1ストッパー 行 異常表示 *)
IF HMI_Message_Request[34] THEN HMI_MessageNo[0] := INT#34; END_IF;
(* Rung 34: 【Y721】A(左側) 位置2ストッパー 異常表示 *)
IF HMI_Message_Request[35] THEN HMI_MessageNo[0] := INT#35; END_IF;

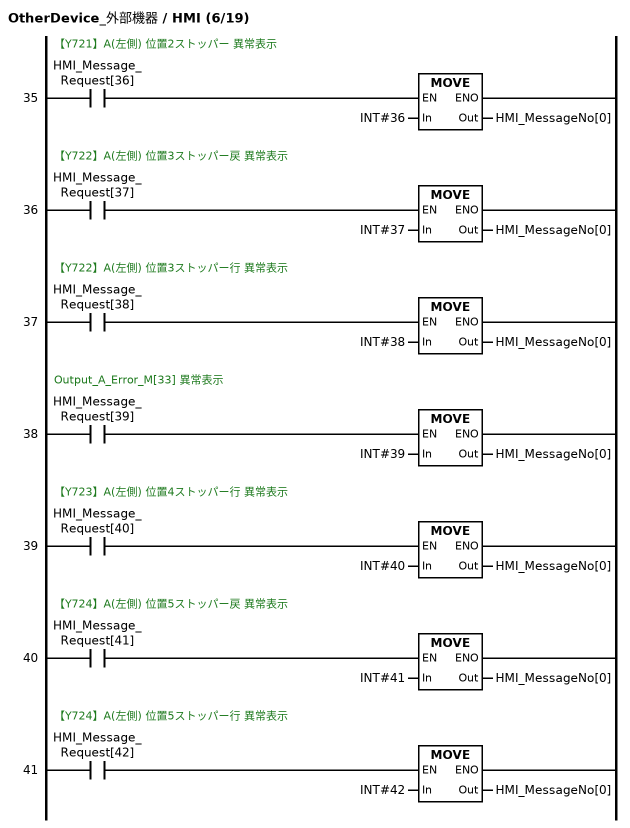
(* Rung 35: 【Y721】A(左側) 位置2ストッパー 異常表示 *)
IF HMI_Message_Request[36] THEN HMI_MessageNo[0] := INT#36; END_IF;
(* Rung 36: 【Y722】A(左側) 位置3ストッパー戻 異常表示 *)
IF HMI_Message_Request[37] THEN HMI_MessageNo[0] := INT#37; END_IF;
(* Rung 37: 【Y722】A(左側) 位置3ストッパー行 異常表示 *)
IF HMI_Message_Request[38] THEN HMI_MessageNo[0] := INT#38; END_IF;
(* Rung 38: Output_A_Error_M[33] 異常表示 *)
IF HMI_Message_Request[39] THEN HMI_MessageNo[0] := INT#39; END_IF;
(* Rung 39: 【Y723】A(左側) 位置4ストッパー行 異常表示 *)
IF HMI_Message_Request[40] THEN HMI_MessageNo[0] := INT#40; END_IF;
(* Rung 40: 【Y724】A(左側) 位置5ストッパー戻 異常表示 *)
IF HMI_Message_Request[41] THEN HMI_MessageNo[0] := INT#41; END_IF;
(* Rung 41: 【Y724】A(左側) 位置5ストッパー行 異常表示 *)
IF HMI_Message_Request[42] THEN HMI_MessageNo[0] := INT#42; END_IF;

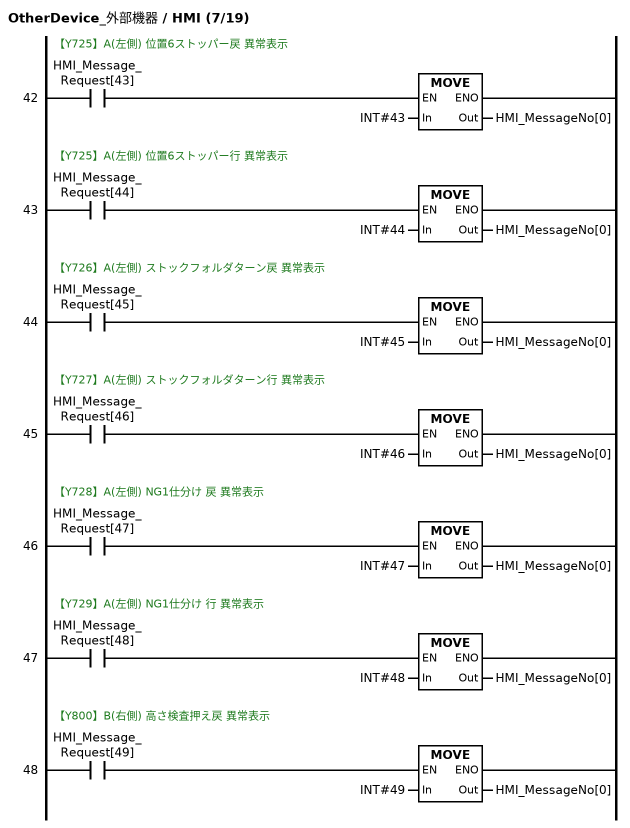
(* Rung 42: 【Y725】A(左側) 位置6ストッパー戻 異常表示 *)
IF HMI_Message_Request[43] THEN HMI_MessageNo[0] := INT#43; END_IF;
(* Rung 43: 【Y725】A(左側) 位置6ストッパー行 異常表示 *)
IF HMI_Message_Request[44] THEN HMI_MessageNo[0] := INT#44; END_IF;
(* Rung 44: 【Y726】A(左側) ストックフォルダターン戻 異常表示 *)
IF HMI_Message_Request[45] THEN HMI_MessageNo[0] := INT#45; END_IF;
(* Rung 45: 【Y727】A(左側) ストックフォルダターン行 異常表示 *)
IF HMI_Message_Request[46] THEN HMI_MessageNo[0] := INT#46; END_IF;
(* Rung 46: 【Y728】A(左側) NG1仕分け 戻 異常表示 *)
IF HMI_Message_Request[47] THEN HMI_MessageNo[0] := INT#47; END_IF;
(* Rung 47: 【Y729】A(左側) NG1仕分け 行 異常表示 *)
IF HMI_Message_Request[48] THEN HMI_MessageNo[0] := INT#48; END_IF;
(* Rung 48: 【Y800】B(右側) 高さ検査押え戻 異常表示 *)
IF HMI_Message_Request[49] THEN HMI_MessageNo[0] := INT#49; END_IF;

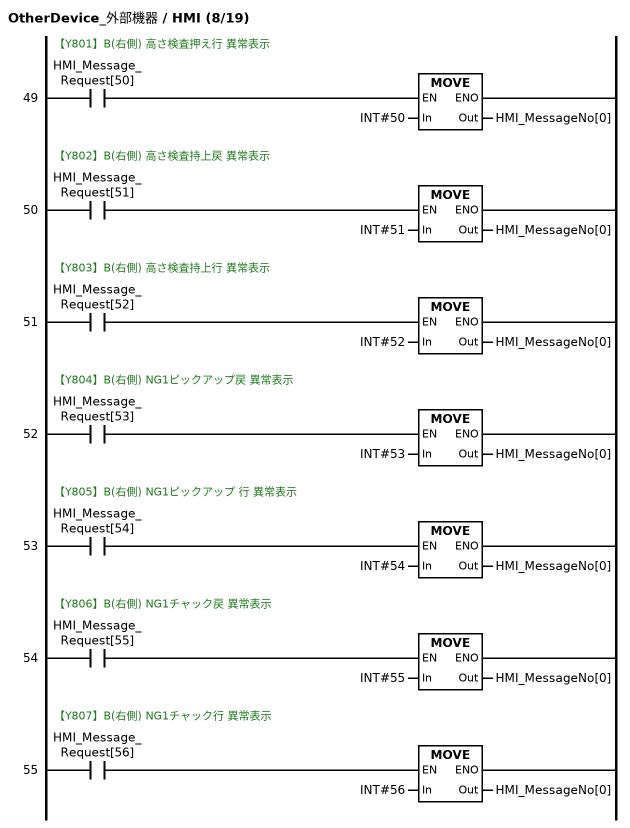
(* Rung 49: 【Y801】B(右側) 高さ検査押え行 異常表示 *)
IF HMI_Message_Request[50] THEN HMI_MessageNo[0] := INT#50; END_IF;
(* Rung 50: 【Y802】B(右側) 高さ検査持上戻 異常表示 *)
IF HMI_Message_Request[51] THEN HMI_MessageNo[0] := INT#51; END_IF;
(* Rung 51: 【Y803】B(右側) 高さ検査持上行 異常表示 *)
IF HMI_Message_Request[52] THEN HMI_MessageNo[0] := INT#52; END_IF;
(* Rung 52: 【Y804】B(右側) NG1ピックアップ戻 異常表示 *)
IF HMI_Message_Request[53] THEN HMI_MessageNo[0] := INT#53; END_IF;
(* Rung 53: 【Y805】B(右側) NG1ピックアップ 行 異常表示 *)
IF HMI_Message_Request[54] THEN HMI_MessageNo[0] := INT#54; END_IF;
(* Rung 54: 【Y806】B(右側) NG1チャック戻 異常表示 *)
IF HMI_Message_Request[55] THEN HMI_MessageNo[0] := INT#55; END_IF;
(* Rung 55: 【Y807】B(右側) NG1チャック行 異常表示 *)
IF HMI_Message_Request[56] THEN HMI_MessageNo[0] := INT#56; END_IF;

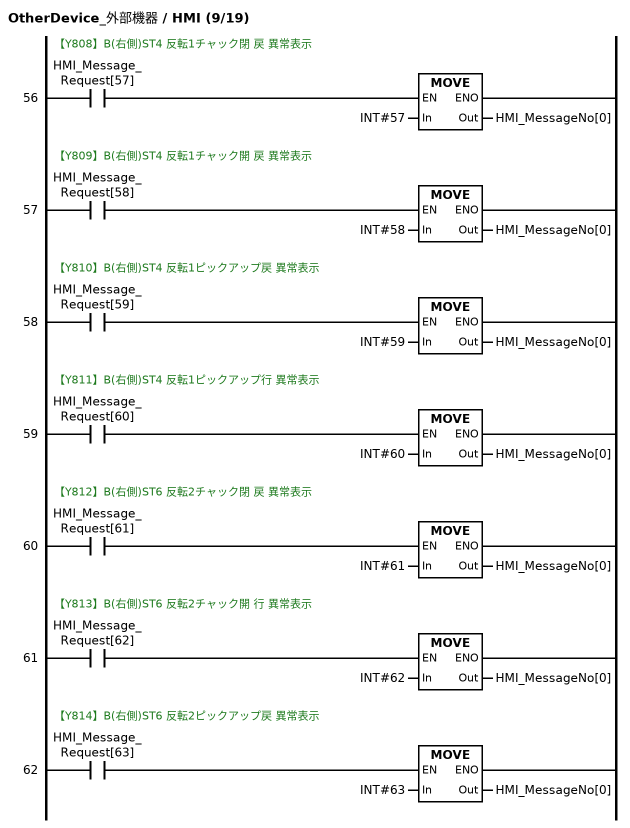
(* Rung 56: 【Y808】B(右側)ST4 反転1チャック閉 戻 異常表示 *)
IF HMI_Message_Request[57] THEN HMI_MessageNo[0] := INT#57; END_IF;
(* Rung 57: 【Y809】B(右側)ST4 反転1チャック開 戻 異常表示 *)
IF HMI_Message_Request[58] THEN HMI_MessageNo[0] := INT#58; END_IF;
(* Rung 58: 【Y810】B(右側)ST4 反転1ピックアップ戻 異常表示 *)
IF HMI_Message_Request[59] THEN HMI_MessageNo[0] := INT#59; END_IF;
(* Rung 59: 【Y811】B(右側)ST4 反転1ピックアップ行 異常表示 *)
IF HMI_Message_Request[60] THEN HMI_MessageNo[0] := INT#60; END_IF;
(* Rung 60: 【Y812】B(右側)ST6 反転2チャック閉 戻 異常表示 *)
IF HMI_Message_Request[61] THEN HMI_MessageNo[0] := INT#61; END_IF;
(* Rung 61: 【Y813】B(右側)ST6 反転2チャック開 行 異常表示 *)
IF HMI_Message_Request[62] THEN HMI_MessageNo[0] := INT#62; END_IF;
(* Rung 62: 【Y814】B(右側)ST6 反転2ピックアップ戻 異常表示 *)
IF HMI_Message_Request[63] THEN HMI_MessageNo[0] := INT#63; END_IF;

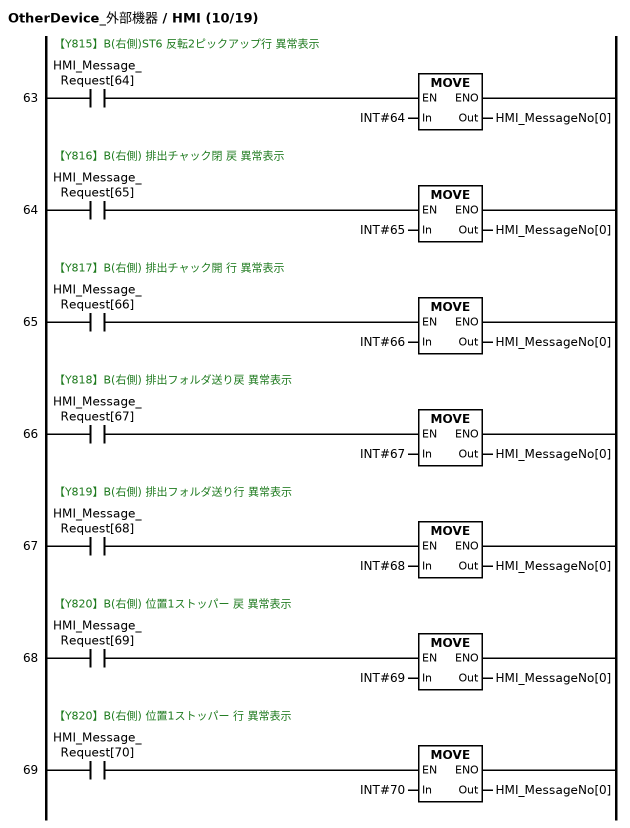
(* Rung 63: 【Y815】B(右側)ST6 反転2ピックアップ行 異常表示 *)
IF HMI_Message_Request[64] THEN HMI_MessageNo[0] := INT#64; END_IF;
(* Rung 64: 【Y816】B(右側) 排出チャック閉 戻 異常表示 *)
IF HMI_Message_Request[65] THEN HMI_MessageNo[0] := INT#65; END_IF;
(* Rung 65: 【Y817】B(右側) 排出チャック開 行 異常表示 *)
IF HMI_Message_Request[66] THEN HMI_MessageNo[0] := INT#66; END_IF;
(* Rung 66: 【Y818】B(右側) 排出フォルダ送り戻 異常表示 *)
IF HMI_Message_Request[67] THEN HMI_MessageNo[0] := INT#67; END_IF;
(* Rung 67: 【Y819】B(右側) 排出フォルダ送り行 異常表示 *)
IF HMI_Message_Request[68] THEN HMI_MessageNo[0] := INT#68; END_IF;
(* Rung 68: 【Y820】B(右側) 位置1ストッパー 戻 異常表示 *)
IF HMI_Message_Request[69] THEN HMI_MessageNo[0] := INT#69; END_IF;
(* Rung 69: 【Y820】B(右側) 位置1ストッパー 行 異常表示 *)
IF HMI_Message_Request[70] THEN HMI_MessageNo[0] := INT#70; END_IF;

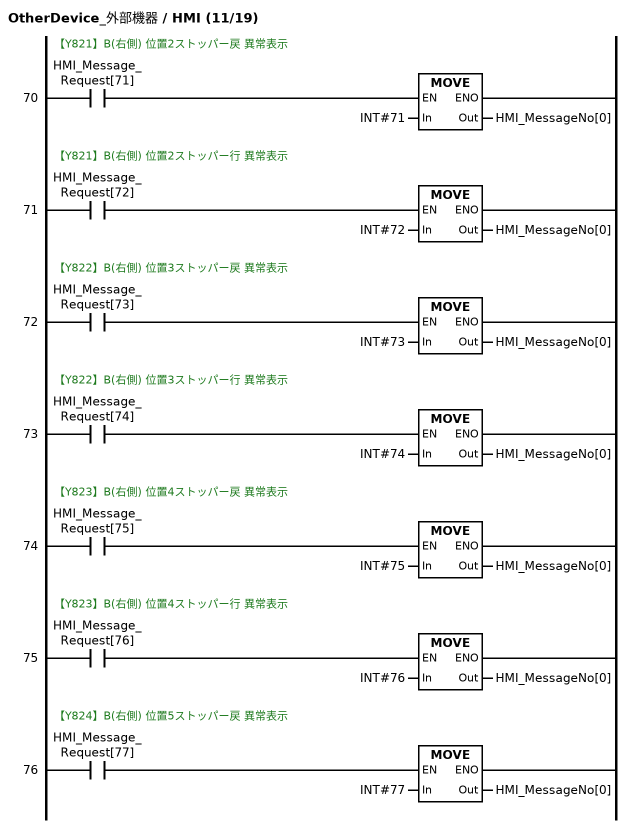
(* Rung 70: 【Y821】B(右側) 位置2ストッパー戻 異常表示 *)
IF HMI_Message_Request[71] THEN HMI_MessageNo[0] := INT#71; END_IF;
(* Rung 71: 【Y821】B(右側) 位置2ストッパー行 異常表示 *)
IF HMI_Message_Request[72] THEN HMI_MessageNo[0] := INT#72; END_IF;
(* Rung 72: 【Y822】B(右側) 位置3ストッパー戻 異常表示 *)
IF HMI_Message_Request[73] THEN HMI_MessageNo[0] := INT#73; END_IF;
(* Rung 73: 【Y822】B(右側) 位置3ストッパー行 異常表示 *)
IF HMI_Message_Request[74] THEN HMI_MessageNo[0] := INT#74; END_IF;
(* Rung 74: 【Y823】B(右側) 位置4ストッパー戻 異常表示 *)
IF HMI_Message_Request[75] THEN HMI_MessageNo[0] := INT#75; END_IF;
(* Rung 75: 【Y823】B(右側) 位置4ストッパー行 異常表示 *)
IF HMI_Message_Request[76] THEN HMI_MessageNo[0] := INT#76; END_IF;
(* Rung 76: 【Y824】B(右側) 位置5ストッパー戻 異常表示 *)
IF HMI_Message_Request[77] THEN HMI_MessageNo[0] := INT#77; END_IF;

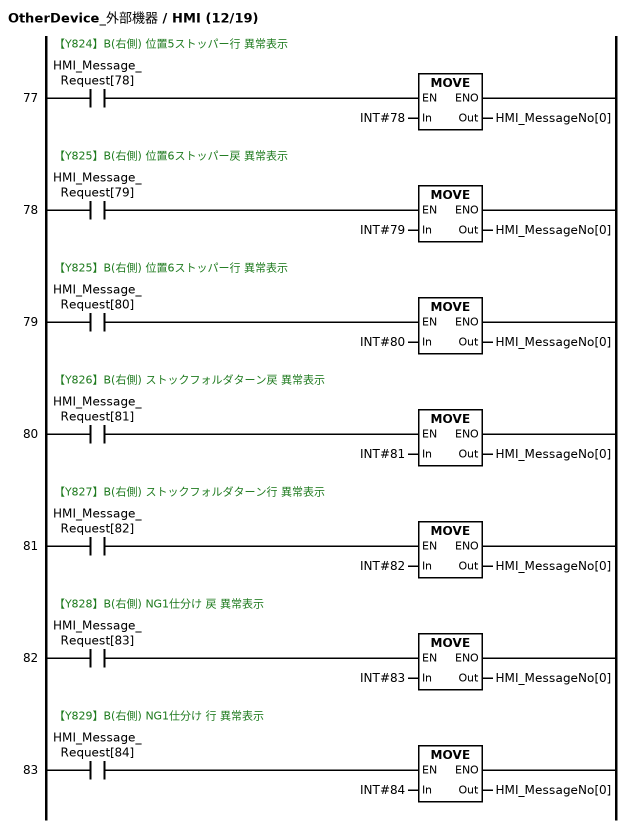
(* Rung 77: 【Y824】B(右側) 位置5ストッパー行 異常表示 *)
IF HMI_Message_Request[78] THEN HMI_MessageNo[0] := INT#78; END_IF;
(* Rung 78: 【Y825】B(右側) 位置6ストッパー戻 異常表示 *)
IF HMI_Message_Request[79] THEN HMI_MessageNo[0] := INT#79; END_IF;
(* Rung 79: 【Y825】B(右側) 位置6ストッパー行 異常表示 *)
IF HMI_Message_Request[80] THEN HMI_MessageNo[0] := INT#80; END_IF;
(* Rung 80: 【Y826】B(右側) ストックフォルダターン戻 異常表示 *)
IF HMI_Message_Request[81] THEN HMI_MessageNo[0] := INT#81; END_IF;
(* Rung 81: 【Y827】B(右側) ストックフォルダターン行 異常表示 *)
IF HMI_Message_Request[82] THEN HMI_MessageNo[0] := INT#82; END_IF;
(* Rung 82: 【Y828】B(右側) NG1仕分け 戻 異常表示 *)
IF HMI_Message_Request[83] THEN HMI_MessageNo[0] := INT#83; END_IF;
(* Rung 83: 【Y829】B(右側) NG1仕分け 行 異常表示 *)
IF HMI_Message_Request[84] THEN HMI_MessageNo[0] := INT#84; END_IF;

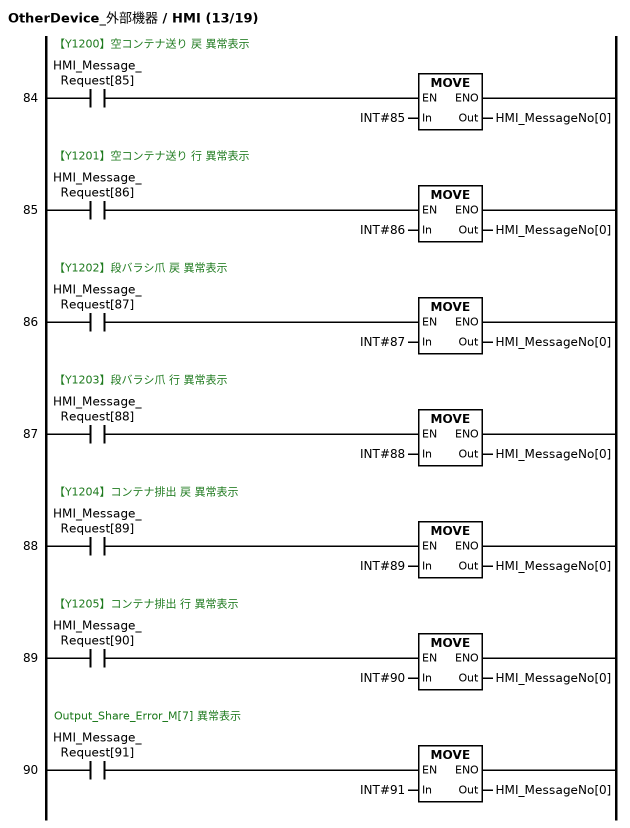
(* Rung 84: 【Y1200】空コンテナ送り 戻 異常表示 *)
IF HMI_Message_Request[85] THEN HMI_MessageNo[0] := INT#85; END_IF;
(* Rung 85: 【Y1201】空コンテナ送り 行 異常表示 *)
IF HMI_Message_Request[86] THEN HMI_MessageNo[0] := INT#86; END_IF;
(* Rung 86: 【Y1202】段バラシ爪 戻 異常表示 *)
IF HMI_Message_Request[87] THEN HMI_MessageNo[0] := INT#87; END_IF;
(* Rung 87: 【Y1203】段バラシ爪 行 異常表示 *)
IF HMI_Message_Request[88] THEN HMI_MessageNo[0] := INT#88; END_IF;
(* Rung 88: 【Y1204】コンテナ排出 戻 異常表示 *)
IF HMI_Message_Request[89] THEN HMI_MessageNo[0] := INT#89; END_IF;
(* Rung 89: 【Y1205】コンテナ排出 行 異常表示 *)
IF HMI_Message_Request[90] THEN HMI_MessageNo[0] := INT#90; END_IF;
(* Rung 90: Output_Share_Error_M[7] 異常表示 *)
IF HMI_Message_Request[91] THEN HMI_MessageNo[0] := INT#91; END_IF;

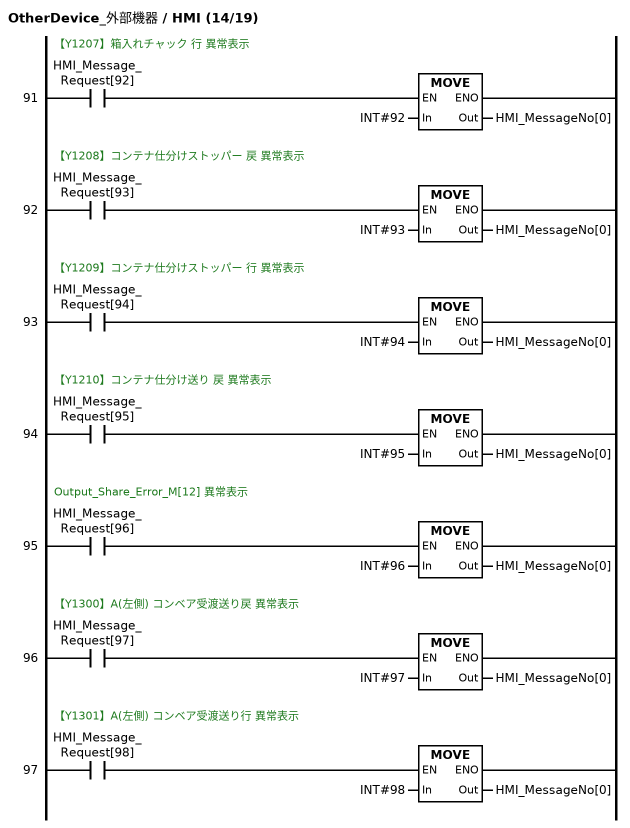
(* Rung 91: 【Y1207】箱入れチャック 行 異常表示 *)
IF HMI_Message_Request[92] THEN HMI_MessageNo[0] := INT#92; END_IF;
(* Rung 92: 【Y1208】コンテナ仕分けストッパー 戻 異常表示 *)
IF HMI_Message_Request[93] THEN HMI_MessageNo[0] := INT#93; END_IF;
(* Rung 93: 【Y1209】コンテナ仕分けストッパー 行 異常表示 *)
IF HMI_Message_Request[94] THEN HMI_MessageNo[0] := INT#94; END_IF;
(* Rung 94: 【Y1210】コンテナ仕分け送り 戻 異常表示 *)
IF HMI_Message_Request[95] THEN HMI_MessageNo[0] := INT#95; END_IF;
(* Rung 95: Output_Share_Error_M[12] 異常表示 *)
IF HMI_Message_Request[96] THEN HMI_MessageNo[0] := INT#96; END_IF;
(* Rung 96: 【Y1300】A(左側) コンベア受渡送り戻 異常表示 *)
IF HMI_Message_Request[97] THEN HMI_MessageNo[0] := INT#97; END_IF;
(* Rung 97: 【Y1301】A(左側) コンベア受渡送り行 異常表示 *)
IF HMI_Message_Request[98] THEN HMI_MessageNo[0] := INT#98; END_IF;

